% RSLogix 500 project L11_CTD.RSS, saved by version 8.30.00.16 %
PROJECT "UNTITLED"    % processor: MicroLogix 1000 %

PROGRAM FILES
  LAD 2 "MAIN_PROG"  7 rungs
  LAD 3 "USER_FAULT"  1 rungs
  LAD 4 "HSC_INT"  1 rungs
  LAD 5 "STI_INT"  1 rungs
  LAD 6, 7, 8, 9, 10, 11, 12, 13, 14, 15, 16: only END

DATA FILES
  O0 OUTPUT  5 elements
  I1 INPUT  8 elements
  S2 STATUS  33 elements
  B3 BINARY  32 elements
  T4 TIMER  40 elements
  C5 COUNTER  32 elements
  R6 CONTROL  16 elements
  N7 INTEGER  105 elements

LADDER 2 "MAIN_PROG"
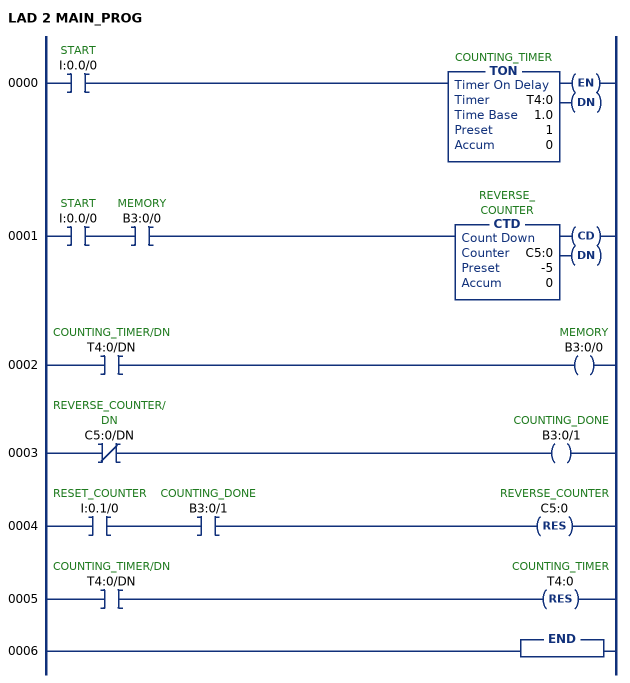
% Rung: 0 %
SOR XIC I:0.0/0 TON T4:0 1.0 1 0 EOR
%   I:0.0/0  START %
%   T4:0  COUNTING_TIMER %
% Rung: 1 %
SOR XIC I:0.0/0 XIC B3:0/0 CTD C5:0 -5 0 EOR
%   I:0.0/0  START %
%   B3:0/0  MEMORY %
%   C5:0  REVERSE_COUNTER %
% Rung: 2 %
SOR XIC T4:0/DN OTE B3:0/0 EOR
%   T4:0  COUNTING_TIMER %
%   B3:0/0  MEMORY %
% Rung: 3 %
SOR XIO C5:0/DN OTE B3:0/1 EOR
%   C5:0  REVERSE_COUNTER %
%   B3:0/1  COUNTING_DONE %
% Rung: 4 %
SOR XIC I:0.1/0 XIC B3:0/1 RES C5:0 EOR
%   I:0.1/0  RESET_COUNTER %
%   B3:0/1  COUNTING_DONE %
%   C5:0  REVERSE_COUNTER %
% Rung: 5 %
SOR XIC T4:0/DN RES T4:0 EOR
%   T4:0  COUNTING_TIMER %
% Rung: 6 %
SOR END EOR

DATA TABLE (non-zero values as saved)
DATA T4
% .PRE .ACC %
% T4:0 % 1 0
DATA C5
% .PRE .ACC %
% C5:0 % -5 0
